(* IEC 61131-3 sources: icsquartz-ndss2025/compiler/libs/wrappers/codesys/SysSocket23, 3 files *)

(* ---- DataTypes.st ---- *)
TYPE INADDR : STRUCT
    S_addr : DWORD;
END_STRUCT
END_TYPE

TYPE SOCKADDRESS : STRUCT
    sin_family : INT;
    sin_port : UINT;
    sin_addr : UDINT;
    sin_zero : ARRAY [0..7] OF SINT;
END_STRUCT
END_TYPE

TYPE SOCKET_FD_SET : STRUCT
    fd_count : UDINT;
    fd_array : ARRAY [0..MAX_SOCKET_FD_SETSIZE] OF DINT;
END_STRUCT
END_TYPE

TYPE SOCKET_LINGER : STRUCT
    l_onoff : WORD;
    l_linger : WORD;
END_STRUCT
END_TYPE

TYPE SOCKET_TIMEVAL : STRUCT
    tv_sec : DINT;
    tv_usec : DINT;
END_STRUCT
END_TYPE

(* ---- GlobalVariables.st ---- *)
VAR_GLOBAL CONSTANT
    SOCKET_INVALID : DINT := -1;
    SOCKET_AF_UNSPEC : INT := 0; (*unspecified*)
    SOCKET_AF_LOCAL : INT := 1; (*local to host (pipes, portals)*)
    SOCKET_AF_UNIX : INT := SOCKET_AF_LOCAL; (*backward compatibility*)
    SOCKET_AF_INET : INT := 2; (*internetwork: UDP, TCP, etc.*)
    SOCKET_AF_IMPLINK : INT := 3; (*arpanet imp addresses*)
    SOCKET_AF_PUP : INT := 4; (*pup protocols: e.g. BSP*)
    SOCKET_AF_CHAOS : INT := 5; (*mit CHAOS protocols*)
    SOCKET_AF_NS : INT := 6; (*XEROX NS protocols*)
    SOCKET_AF_ISO : INT := 7; (*ISO protocols*)
    SOCKET_AF_OSI : INT := SOCKET_AF_ISO;
    SOCKET_AF_ECMA : INT := 8; (*european computer manufacturers*)
    SOCKET_AF_DATAKIT : INT := 9; (*datakit protocols*)
    SOCKET_AF_CCITT : INT := 10; (*CCITT protocols, X.25 etc*)
    SOCKET_AF_SNA : INT := 11; (*IBM SNA*)
    SOCKET_AF_DECnet : INT := 12; (*DECnet*)
    SOCKET_AF_DLI : INT := 13; (*DEC Direct data link interface*)
    SOCKET_AF_LAT : INT := 14; (*LAT*)
    SOCKET_AF_HYLINK : INT := 15; (*NSC Hyperchannel*)
    SOCKET_AF_APPLETALK : INT := 16; (*Apple Talk*)
    SOCKET_AF_ROUTE : INT := 17; (*Internal Routing Protocol*)
    SOCKET_AF_LINK : INT := 18; (*Link layer interface*)
    SOCKET_pseudo_AF_XTP : INT := 19; (*eXpress Transfer Protocol (no AF)*)
    SOCKET_AF_COIP : INT := 20; (*connection-oriented IP, aka ST II*)
    SOCKET_AF_CNT : INT := 21; (*Computer Network Technology*)
    SOCKET_pseudo_AF_RTIP : INT := 22; (*Help Identify RTIP packets*)
    SOCKET_AF_IPX : INT := 23; (*Novell Internet Protocol*)
    SOCKET_AF_SIP : INT := 24; (*Simple Internet Protocol*)
    SOCKET_pseudo_AF_PIP : INT := 25; (*Help Identify PIP packets*)
    SOCKET_AF_MAX : INT := 26;
    SOCKET_AF_INET_BSD : INT := 100; (*BSD-specific INET af*)
    SOCKET_AF_INET_STREAMS : INT := 101; (*STREAMS-specific INET af*)
    SOCKET_SOL : WORD := 16#FFFF; (*Level number for (get/set)sockopt() to apply to socket itself.*)
    SOCKET_SO_DEBUG : DINT := 16#1; (*turn on debugging info recording*)
    SOCKET_SO_ACCEPTCONN : DINT := 16#2; (*socket has had listen()*)
    SOCKET_SO_REUSEADDR : DINT := 16#4; (*allow local address reuse*)
    SOCKET_SO_KEEPALIVE : DINT := 16#8; (*keep connections alive*)
    SOCKET_SO_DONTROUTE : DINT := 16#10; (*just use interface addresses*)
    SOCKET_SO_BROADCAST : DINT := 16#20; (*permit sending of broadcast msgs*)
    SOCKET_SO_USELOOPBACK : DINT := 16#40; (*bypass hardware when possible*)
    SOCKET_SO_LINGER : DINT := 16#80; (*linger on close if data present*)
    SOCKET_SO_OOBINLINE : DINT := 16#100; (*leave received OOB data in line*)
    SOCKET_SO_REUSEPORT : DINT := 16#200; (*allow local address & port reuse*)
    SOCKET_SO_SNDBUF : DINT := 16#1001; (*send buffer size*)
    SOCKET_SO_RCVBUF : DINT := 16#1002; (*receive buffer size*)
    SOCKET_SO_SNDLOWAT : DINT := 16#1003; (*send low-water mark*)
    SOCKET_SO_RCVLOWAT : DINT := 16#1004; (*receive low-water mark*)
    SOCKET_SO_SNDTIMEO : DINT := 16#1005; (*send timeout*)
    SOCKET_SO_RCVTIMEO : DINT := 16#1006; (*receive timeout*)
    SOCKET_SO_ERROR : DINT := 16#1007; (*get error status and clear*)
    SOCKET_SO_TYPE : DINT := 16#1008; (*get socket type*)
    SOCKET_SO_PROTOTYPE : DINT := 16#1009; (*get/set protocol type*)
    SOCKET_TCP_NODELAY : DINT := 16#1; (*don’t delay send to coalesce packets*)
    SOCKET_TCP_MAXSEG : DINT := 16#2; (*set maximum segment size*)
    SOCKET_STREAM : DINT := 1; (*stream socket*)
    SOCKET_DGRAM : DINT := 2; (*datagram socket*)
    SOCKET_RAW : DINT := 3; (*raw-protocol interface*)
    SOCKET_RDM : DINT := 4; (*reliably-delivered message*)
    SOCKET_SEQPACKET : DINT := 5; (*sequenced packet stream*)
    SOCKET_INADDR_ANY : UDINT := 16#0; (*Inet address definitions*)
    SOCKET_INADDR_LOOPBACK : UDINT := 16#7F000001;
    SOCKET_INADDR_BROADCAST : UDINT := 16#FFFFFFFF;
    SOCKET_INADDR_NONE : UDINT := 16#FFFFFFFF;
    SOCKET_IPPROTO_IP : DINT := 0; (*dummy for IP*)
    SOCKET_IPPROTO_ICMP : DINT := 1; (*control message protocol*)
    SOCKET_IPPROTO_IGMP : DINT := 2; (*group management protocol*)
    SOCKET_IPPROTO_GGP : DINT := 3; (*gateway^2 (deprecated)*)
    SOCKET_IPPROTO_TCP : DINT := 6; (*tcp*)
    SOCKET_IPPROTO_PUP : DINT := 12; (*pup*)
    SOCKET_IPPROTO_UDP : DINT := 17; (*user datagram protocol*)
    SOCKET_IPPROTO_IDP : DINT := 22; (*xns idp*)
    SOCKET_IPPROTO_ND : DINT := 77; (*UNOFFICIAL net disk proto*)
    SOCKET_IPPROTO_RAW : DINT := 255; (*raw IP packet*)
    SOCKET_IPPROTO_MAX : DINT := 256;
    SOCKET_MSG_OOB : DINT := 16#1; (*process out-of-band data*)
    SOCKET_MSG_PEEK : DINT := 16#2; (*peek at incoming message*)
    SOCKET_MSG_DONTROUTE : DINT := 16#4; (*send without using routing tables*)
    SOCKET_FIONREAD : DINT := 1; (*get num chars available to read*)
    SOCKET_FIONBIO : DINT := 2; (*set to non-blocking*)
    SOCKET_FD_SETSIZE : DINT := 64; (*For SysSockSelect() descriptors*)
    MAX_SOCKET_FD_SETSIZE : DINT := 63;
END_VAR

(* ---- POUs.st ---- *)
FUNCTION SysSockAccept : DINT
VAR_INPUT
    diSocket : DINT;
    pSockAddr : DWORD;  // Address of SocketAddress (SOCKADDRESS)
    piSockAddrSize : DWORD;  // Address of socket address size (DINT)
END_VAR

unimplemented('SysSockAccept');
END_FUNCTION

FUNCTION SysSockBind : BOOL
VAR_INPUT
    diSocket : DINT;
    pSockAddr : DWORD;  // Address of SocketAddress (SOCKADDRESS)
    diSockAddrSize : DINT;  // Size of socket address
END_VAR

unimplemented('SysSockBind');
END_FUNCTION

FUNCTION SysSockClose : BOOL
VAR_INPUT
    diSocket : DINT;
END_VAR

unimplemented('SysSockClose');
END_FUNCTION

FUNCTION SysSockConnect : BOOL
VAR_INPUT
    diSocket : DINT;
    pSockAddr : DWORD;  // Address of SocketAddress (SOCKADDRESS)
    diSockAddrSize : DINT;  // Size of socket address
END_VAR

unimplemented('SysSockConnect');
END_FUNCTION

FUNCTION SysSockCreate : DINT
VAR_INPUT
    diAddressFamily : DINT;
    diType : DINT;
    diProtocol : DINT;
END_VAR

unimplemented('SysSockCreate');
END_FUNCTION

FUNCTION SysSockGetHostByName : DWORD
VAR_INPUT
    stHostName : STRING;
END_VAR

unimplemented('SysSockGetHostByName');
END_FUNCTION

FUNCTION SysSockGetHostName : BOOL
VAR_INPUT
    diNameLength : DINT;
END_VAR
VAR_IN_OUT
    stHostName : STRING;
END_VAR

unimplemented('SysSockGetHostName');
END_FUNCTION

FUNCTION_BLOCK SysSockGetLastError
VAR_INPUT
    bEnable : BOOL;
    diSocket : DINT;
END_VAR
VAR_OUTPUT
    bDone : BOOL;
    bBusy : BOOL;
    bError : BOOL;
    wErrorId : WORD;
    dwLastError : DWORD;
END_VAR

unimplemented('SysSockGetLastError');
END_FUNCTION_BLOCK

FUNCTION SysSockGetLastErrorSync : DINT
VAR_INPUT
    diSocket : DINT;
END_VAR

unimplemented('SysSockGetLastErrorSync');
END_FUNCTION

FUNCTION SysSockGetOption : BOOL
VAR_INPUT
    diSocket : DINT;
    diLevel : DINT;
    diOption : DINT;
    pOptionValue : DWORD;    // Address of option
    piOptionLength : DWORD;  // Address of option size (DINT)
END_VAR

unimplemented('SysSockGetOption');
END_FUNCTION

FUNCTION SysSockHtonl : DWORD
VAR_INPUT
    dwHost : DWORD;
END_VAR

unimplemented('SysSockHtonl');
END_FUNCTION

FUNCTION SysSockHtons : WORD
VAR_INPUT
    wHost : WORD;
END_VAR

unimplemented('SysSockHtons');
END_FUNCTION

FUNCTION SysSockInetAddr : DWORD
VAR_IN_OUT
    stIPAddr : STRING;
END_VAR

unimplemented('SysSockInetAddr');
END_FUNCTION

FUNCTION SysSockInetNtoa : BOOL
VAR_INPUT
    InAddr : INADDR;
    diIPAddrSize : DINT;
END_VAR
VAR_IN_OUT
    stIPAddr : STRING;
END_VAR

unimplemented('SysSockInetNtoa');
END_FUNCTION

FUNCTION SysSockIoctl : DINT
VAR_INPUT
    diSocket : DINT;
    diCommand : DINT;
    piParameter : DWORD; // Address of parameter (DINT)
END_VAR

unimplemented('SysSockIoctl');
END_FUNCTION

FUNCTION SysSockListen : BOOL
VAR_INPUT
    diSocket : DINT;
    diMaxConnections : DINT;
END_VAR

unimplemented('SysSockListen');
END_FUNCTION

FUNCTION SysSockNtohl : DWORD
VAR_INPUT
    dwNet : DWORD;
END_VAR

unimplemented('SysSockNtohl');
END_FUNCTION

FUNCTION SysSockNtohs : WORD
VAR_INPUT
    wNet : WORD;
END_VAR

unimplemented('SysSockNtohs');
END_FUNCTION

FUNCTION SysSockSelect : DINT
VAR_INPUT
    diWidth : DINT;        // Typically SOCKET_FD_SETSIZE
    fdRead : DWORD;        // Address of SOCKET_FD_SET
    fdWrite : DWORD;       // Address of SOCKET_FD_SET
    fdExcept : DWORD;      // Address of SOCKET_FD_SET
    ptvTimeout : DWORD;    // Address of SOCKET_TIMEVAL
END_VAR

// This routine permits a task to pend until one of a set of sockets handles becomes ready.
// Three parameters – fdRead, fdWrite and fdExcept – point to file descriptor sets in which each array entry corresponds to a particular socket handle.
// If a socket handle is not ready, it will be written in the array to -1 (SOCKET_INVALID).
// With the timeout value, a timeout for the operation can be specified. diWidth is the size of the fd_array array in SOCKETFD_SET.
// The function returns the operating system result.
// <0: Error 0: Timeout expired >0: Typically number of sockets that are successfully selected
unimplemented('SysSockSelect');
END_FUNCTION

FUNCTION SysSockSetIPAddress : BOOL
VAR_INPUT
    stCardName : STRING;     // Card Name
    stIPAddress : STRING;    // IP Address
END_VAR

unimplemented('SysSockSetIPAddress');
END_FUNCTION

FUNCTION SysSockSetOption : BOOL
VAR_INPUT
    diSocket : DINT;            // Socket
    diLevel : DINT;             // Level
    diOption : DINT;            // Option
    pOptionValue : DWORD;       // Address of option
    diOptionLength : DINT;      // Length of option
END_VAR

unimplemented('SysSockSetOption');
END_FUNCTION

FUNCTION SysSockShutdown : BOOL
VAR_INPUT
    diSocket : DINT;   // Socket
    diHow : DINT;      // How
END_VAR

unimplemented('SysSockShutdown');
END_FUNCTION

FUNCTION SysSockRecv : DINT
VAR_INPUT
    diSocket : DINT;         // Socket
    pbyBuffer : DWORD;       // Address of buffer to receive
    diBufferSize : DINT;     // Buffer Size
    diFlags : DINT;          // Flags
END_VAR

unimplemented('SysSockRecv');
END_FUNCTION

FUNCTION SysSockSend : DINT
VAR_INPUT
    diSocket : DINT;         // Socket
    pbyBuffer : DWORD;       // Address of buffer to send
    diBufferSize : DINT;     // Buffer Size
    diFlags : DINT;          // Flags
END_VAR

unimplemented('SysSockSend');
END_FUNCTION

FUNCTION SysSockRecvFrom : DINT
VAR_INPUT
    diSocket : DINT;         // Socket
    pbyBuffer : DWORD;       // Address of buffer to receive
    diBufferSize : DINT;     // Buffer Size
    diFlags : DINT;          // Flags
    pSockAddr : DWORD;       // Address of socket address SOCKADDRESS
    diSockAddrSize : DINT;   // Size of socket address
END_VAR

unimplemented('SysSockRecvFrom');
END_FUNCTION

FUNCTION SysSockSendTo : DINT
VAR_INPUT
    diSocket : DINT;         // Socket
    pbyBuffer : DWORD;       // Address of buffer to receive
    diBufferSize : DINT;     // Buffer Size
    diFlags : DINT;          // Flags
    pSockAddr : DWORD;       // Address of socket address SOCKADDRESS
    diSockAddrSize : DINT;   // Size of socket address
END_VAR

unimplemented('SysSockSendTo');
END_FUNCTION
